Fanuc TP program (LS listing): PickWindsh.LS

/PROG  PickWindsh
/ATTR
OWNER		= MNEDITOR;
COMMENT		= "RoboDK sequence";
PROG_SIZE	= 0;
CREATE		= DATE 31-12-14  TIME 12:00:00;
MODIFIED	= DATE 31-12-14  TIME 12:00:00;
FILE_NAME	= PickWindsh;
VERSION		= 0;
LINE_COUNT	= 24;
MEMORY_SIZE	= 0;
PROTECT		= READ_WRITE;
TCD:  STACK_SIZE	= 0,
      TASK_PRIORITY	= 50,
      TIME_SLICE	= 0,
      BUSY_LAMP_OFF	= 0,
      ABORT_REQUEST	= 0,
      PAUSE_REQUEST	= 0;
DEFAULT_GROUP	= 1,*,*,*,*,*,*;
CONTROL_CODE	= 00000000 00000000;
/MN
   1:  ! Program generated by VerticalBot Studio for Fanuc M-710iC/45M ;
   2:  ! on 25/10/2026 12:00:00 ;
   3:  ! Using nominal kinematics. ;
   4:  PR[9,1]=2299.810 ;
   5:  PR[9,2]=1718.890 ;
   6:  PR[9,3]=-421.206 ;
   7:  PR[9,4]=0.000 ;
   8:  PR[9,5]=0.000 ;
   9:  PR[9,6]=-180.000 ;
  10:  UFRAME[9]=PR[9] ;
  11:  UFRAME_NUM=9 ;
  12:  PR[9,1]=0.000 ;
  13:  PR[9,2]=0.000 ;
  14:  PR[9,3]=110.022 ;
  15:  PR[9,4]=0.000 ;
  16:  PR[9,5]=0.000 ;
  17:  PR[9,6]=0.000 ;
  18:  UTOOL[9]=PR[9] ;
  19:  UTOOL_NUM=9 ;
  20:J P[1] 20% FINE ;
  21:L P[2] 200mm/sec FINE ;
  22:  ! Attach to Tool Windshield ;
  23:  WAIT  0.25(sec) ;
  24:L P[3] 200mm/sec FINE ;
/POS
P[1]{
   GP1:
    UF : 9, UT : 9,
	J1=    45.094 deg,	J2=    34.535 deg,	J3=    -59.541 deg,
	J4=    -49.332 deg,	J5=    69.031 deg,	J6=    22.613 deg
};
P[2]{
   GP1:
    UF : 9, UT : 9,        CONFIG : 'N U T, 0, 0, 0',
	X =   459.506  mm,	Y =   582.163  mm,	Z =   338.451  mm,
	W =     0.000 deg,	P =   -90.000 deg,	R =     0.000 deg
};
P[3]{
   GP1:
    UF : 9, UT : 9,        CONFIG : 'N U B, 0, 0, -1',
	X =   458.000  mm,	Y =   582.163  mm,	Z =  1000.000  mm,
	W =     0.000 deg,	P =   -90.000 deg,	R =     0.000 deg
};
/END
